FUNCTION_BLOCK ThisXTS EXTENDS Xts<1,1,1>
VAR
	_homePosition : LREAL;
END_VAR

PROPERTY HomePosition : LREAL
GET
HomePosition := _homePosition;
END_GET
SET
_homePosition := HomePosition;
END_SET
END_PROPERTY

METHOD MoverHomeSequence : BOOL
VAR
	i : INT;
END_VAR
FOR i := 0 TO _registeredNumberOfMovers - 1 DO 
	iMovers[i].MoveTo(_homePosition,1000.0,FALSE);
END_FOR
END_METHOD

END_FUNCTION_BLOCK

(* stored: Version 1.1.0.1, ProductVersion 3.1.4026.21
   POU ThisXTS: Id {adc628a7-7a2e-4111-937d-b66eb159493c}, SpecialFunc None
   Property HomePosition: Id {d602f7c2-50bd-47cc-89fa-7135c8d1eaba}
   Get Get: Id {86043ce9-0793-47f3-b3e8-793e99e740e9}
   Set Set: Id {56cccc03-60ff-4ea7-9531-591ff5482e5e}
   Method MoverHomeSequence: Id {dd65f3ed-d01b-4f9f-95cc-8438905256ec} *)
